Fanuc KAREL source: kt00118.KL

-- PROVISIONAL review KL for V1013-1; original PC SHA256 8e96ca13d22c23ca25408edeb8b6b089b044299d3efb354f7c4e56db8bcb911a
-- Incomplete behavior may be omitted. Consult companion uncertainty JSON. Do not deploy.
PROGRAM KT00118
%NOLOCKGROUP
VAR
  OUT : REAL
-- UNRESOLVED_DECL Y1 type=002018
-- UNRESOLVED_DECL Y2 type=002018
BEGIN
  -- UNRESOLVED_PC offsets 5-19; opcodes 2E,22,9D,33,B2
  -- UNRESOLVED_PC offsets 24-38; opcodes 2E,22,9D,33,B2
  -- UNRESOLVED_PC offsets 43-57; opcodes 2E,22,9D,33,B2
  -- UNRESOLVED_PC offsets 62-76; opcodes 2E,22,9D,33,B2
  -- UNRESOLVED_PC offsets 81-110; opcodes 22,9D,33,B1,22,9D,33,B1,64,29,64,29,6C,23
  -- UNRESOLVED_PC offsets 115-119; opcodes 7F
END KT00118
